(*
SPDX-FileCopyrightText: © 2026 Oleksandr Tiutyk <trofimich@gmail.com>
SPDX-License-Identifier: MIT
License: https://opensource.org/license/mit
*)

(*!
<summary>Runs one workflow contract scenario in an isolated fixture.</summary>
<description>
Owns a freshly allocated fixture for the active run. AfterTest releases it after success or a reported
exception. A concrete pointer preserves FB_exit for the fixture and its nested resource owners.
Use one task. Do not copy the test case while it owns a fixture.
</description>
*)

{attribute 'no_assign'}
{attribute 'no_explicit_call' := 'do not call this function block directly'}
FUNCTION_BLOCK WorkflowContractTestCase EXTENDS TOF_Testing.SingleCycleTest
VAR_STAT
	{attribute 'hide'}
	_ClassName : STRING := __POUNAME();
END_VAR
VAR
	_Scenario : WORKFLOW_CONTRACT_TEST_SCENARIO;
	_Fixture : POINTER TO WorkflowContractTestFixture;
END_VAR

(*!
<summary>Selects the scenario without allocating its fixture.</summary>
<param name="name">Name reported for this case.</param>
<param name="parent">Group that owns this case.</param>
<param name="scenario">Scenario selected for the case.</param>
*)
METHOD FB_init : BOOL
VAR_INPUT
	bInitRetains: BOOL; // TRUE: the retain variables are initialized (reset warm / reset cold)
	bInCopyCode: BOOL; // TRUE: the instance will be copied to the copy code afterward (online change)
	name : WSTRING;
	parent : TOF_Testing.ITestElement;
	scenario : WORKFLOW_CONTRACT_TEST_SCENARIO;
END_VAR
IF NOT bInCopyCode THEN
	_Scenario := scenario;
END_IF

FB_init := TRUE;
END_METHOD

(*!
<summary>Allocates a fresh fixture and runs the selected scenario.</summary>
<description>Terminal allocation failure is raised at the task boundary after case handling.</description>
*)
METHOD PROTECTED ExecuteTest
VAR
	assertions : REFERENCE TO TOF_Testing.Assertions;
END_VAR
_Fixture := __NEW(WorkflowContractTestFixture);

IF _Fixture = 0 THEN
	TOF_Core.DynamicMemoryManager.RaiseAllocationFailure();

	RETURN;
END_IF

assertions REF= Assert;
_Fixture^.ExecuteScenario(scenario := _Scenario, assertions := assertions);
END_METHOD

(*!
<summary>Releases the fixture before the case outcome is published.</summary>
<description>The framework records an exception from teardown. Clear the stored alias before releasing.</description>
*)
METHOD PROTECTED AfterTest
VAR
	fixture : POINTER TO WorkflowContractTestFixture;
	released : BOOL;
END_VAR
fixture := _Fixture;
_Fixture := 0;

IF fixture <> 0 THEN
	released := fixture^.TryReleaseLoadedWorkflow();
	__DELETE(fixture);

	IF NOT released THEN
		IF Outcome = TOF_Testing.TEST_OUTCOME.FAILED THEN
			Tc2_System.ADSLOGSTR(
				msgCtrlMask := Tc2_System.Global_Variables.ADSLOG_MSGTYPE_ERROR,
				msgFmtStr := 'Unable to release loaded workflow in %s',
				strArg := TO_STRING(Name)
			);
		ELSE
			RecordFailure(message := "Unable to release loaded workflow");
		END_IF
	END_IF
END_IF
END_METHOD

(*!
<summary>Releases an active fixture if the case is unloaded before its teardown.</summary>
<description>The fixture and its nested FB_exit paths complete without exceptions.</description>
<param name="bInCopyCode">TwinCAT copy-code exit marker. The previous instance leaves copied storage alive.</param>
*)
METHOD FB_exit : BOOL
VAR_INPUT
	bInCopyCode : BOOL;
END_VAR
IF NOT bInCopyCode AND_THEN _Fixture <> 0 THEN
	__DELETE(_Fixture);
END_IF

FB_exit := TRUE;
END_METHOD

(*!
<summary>Borrows the concrete class name. Callers must not modify it.</summary>
*)
{attribute 'monitoring' := 'call'}
PROPERTY ClassName : REFERENCE TO STRING
GET
ClassName REF= _ClassName;
END_GET
END_PROPERTY

(*!
<summary>Borrows the project namespace name. Callers must not modify it.</summary>
*)
{attribute 'monitoring' := 'call'}
PROPERTY NamespaceName : REFERENCE TO STRING
GET
NamespaceName REF= CurrentNamespace.Name;
END_GET
END_PROPERTY

(*!
<summary>Reports the complete instance size in bytes.</summary>
*)
{attribute 'monitoring' := 'call'}
PROPERTY SelfSize : ULINT
GET
SelfSize := XSIZEOF(THIS^);
END_GET
END_PROPERTY

END_FUNCTION_BLOCK

(* stored: Version 1.1.0.1
   POU WorkflowContractTestCase: Id {a9805011-9553-4648-8b05-2eaaf2ddbf8a}, SpecialFunc None
   Method FB_init: Id {9146b617-a2a7-4f45-95c9-bfdd47adcecc}
   Method ExecuteTest: Id {48ac0298-3897-4b94-b6fe-b13f6e655c44}
   Method AfterTest: Id {6e572add-4424-42f2-b9f6-cec8e1d72e94}
   Method FB_exit: Id {d8a5654c-2d07-4f02-a7fe-b2b5875fef04}
   Property ClassName: Id {328da49d-8149-4720-8732-fd346bf92ba7}
   Get Get: Id {78a65a5e-2ced-48f4-92f3-5956dbd96e1e}
   Property NamespaceName: Id {db80ad18-9a5a-4f2e-9f8e-680dd3ad375e}
   Get Get: Id {9a23cc24-cf38-4879-a699-a661cc70b96f}
   Property SelfSize: Id {64943f36-9b40-4817-aaaa-cad6841554fc}
   Get Get: Id {a087ab06-2409-4eb0-8d70-248cb6d890ef} *)
